(* IEC 61131-3 sources: Test002/ConveyorBelt/Class/SafetyBaseFSoE (part 5) *)

    end_if;

    //write to hardware from other module received SDO
    if ( ui_cnt_SDOInputBuffer > 0 ) & p_SDOInputBuffer then

      //set pointer to first SDO in the SDO list
      p_SDO_act   := p_SDOInputBuffer$^SDOHeader;

      //calculate length of SDO (CRC + data length)
      us_SDO_length := sizeof (SDOHeader.StdHeader.CRC) + p_SDO_act^.StdHeader.Len;

      //check, if buffer is empty
      if ( p_Handle_SDO_Write^.us_Status = SAFETY_SDO_NO_DATA ) then

#ifdef SAFETY_PROTOCOL_ANALYZER_ACTIVATED
  RecordFrame(p_SDO_act$^DINT, 1);
#endif

        //copy SDO into write-buffer
        ToStdLib.MemCpy(dest := #p_Handle_SDO_Write^.SDOStructure, source := p_SDO_act, size := us_SDO_length);

        //mark SDO data as valid
        p_Handle_SDO_Write^.us_Status := SAFETY_SDO_DATA_VALID;

        //decrement amount of SDOs
        ui_cnt_SDOInputBuffer -= 1;

        //if there is at least 1 SDO left, copy the remaining memory over the actual SDO
        if ( ui_cnt_SDOInputBuffer > 0 ) then

          //remove first entry in the SDO list
          _memmove(p_SDOInputBuffer, (p_SDOInputBuffer + SBF_SDO_MAX_LENGTH), (ui_cnt_SDOInputBuffer * SBF_SDO_MAX_LENGTH));
        end_if;
      end_if;
    end_if;

    if (b_ManagerInitialisationFinished = TRUE) & ( SafetyState <> _ReinitConfig ) & ( p_Handle_SDO_Write^.us_Status = SAFETY_SDO_NO_DATA ) then

      // priority request before checking the scheduler
      // if the channel is free and we have a command request for the flexible constellation node => send the command
      if (LastRequest = _NoOpenRequest) & (sFlexCon.FoundNodeInConfig) & (sFlexCon.CommandRequest) then

        StandardRequest.SDOHeader.CRC  := 0;                               // CRC is always 0 in Std communication
        StandardRequest.SDOHeader.Cmd  := SBF_SDO_COMMAND_WRITE;           // read command
        StandardRequest.SDOHeader.Typ  := SDO_STD;                         // standard frame type
        StandardRequest.SDOHeader.SeqNr:= StandardSeqNr OR 16#80;          // sequence number
        StandardRequest.SDOHeader.Len  := 4 + 4 + 1 + sizeof(UDINT);       // header + destination address + length of data + size of data
        StandardRequest.aData[0]$UDINT := SBF_SDO_ADDRESS_FLEX_CON_NODE;   // address of the flex con data
        StandardRequest.aData[4]       := sizeof(UDINT);                   // length of data
        StandardRequest.aData[5]$UDINT := sFlexCon.CommandRequest;     // new command

        // reset marker to detect new commands
        sFlexCon.CommandRequest := 0;

        LastRequest := _WriteFlexConCommand;

        //copy SDO into write-buffer
        ToStdLib.MemCpy(dest := #p_Handle_SDO_Write^.SDOStructure, source := #StandardRequest, size := (sizeof(SDOHeader.StdHeader.CRC) + StandardRequest.SDOHeader.Len));

        //mark SDO data as valid
        p_Handle_SDO_Write^.us_Status := SAFETY_SDO_DATA_VALID;

        if ( pISafety^.udVersion >= 16#1001 ) then
          SAFETY_iPushSafetyTask();
        end_if;

      end_if;

      // Start of scheduler; we need to share the time between reading, writing and diagnosis
      us_UnsafeSchedulerRun := 0;

      // number of steps in total minus 1, because the SetBusReady doesn't count here since it's not part of the rotation
      SchedulerStepNo := 10;

      // Check actions until we find somthing we need to do
      // all x (SchedulerStepNo) action-steps must be walked through during one cycle to make sure new data is fetched as fast as possible
      // SetBusReady is an exception: this step is only performed once on bootup!
      while (us_UnsafeSchedulerRun < SchedulerStepNo) & (LastRequest = _NoOpenRequest) do
        us_UnsafeSchedulerRun += 1;
        ud_UnsafeTimeoutCounter := 0; //No active request: we can reset the timeout-counter
        case UnsafeScheduler of
//**********************************************************************************************************************************************************
          UnsafeSchedulerSetBusReady:  // this step is excluded from the rotation (set at startup, on disconnect or quit error)

            case us_SetBusReadyState of

            //-------------------------------------------------------------------------------------------------------------
              WaitPDOsSyncron:

                EverythingSynchron := TRUE;

                // it's possible that all PDOs are coming from a different domain, then we have no inputbuffer
                if ui_cnt_PDOInputBuffer then
                  p_PDOInBufferAct := #aPDOInputBuffer[0];
                  for i := 0 to (ui_cnt_PDOInputBuffer-1) do
                    if p_PDOInBufferAct^.b_TimeSynchron = FALSE then
                      // we're still not synchron with this module. if it's optional it is probably not connected
                      if p_PDOInBufferAct^.b_IsOptional then
                        if (ops.tAbsolute - ud_OptionalTimeoutStart) <= SBF_OPTIONAL_MODULE_SYNC_TIMEOUT then
                          // if timeout not exceeded => not sychron (otherwise the variable will stay on it's old value)
                          EverythingSynchron := FALSE;
                          exit;
                        else
                          TRACE("Synchronisation timeout for optional module exceeded => assume it's synchon.");
                        end_if;
                      else
                        EverythingSynchron := FALSE;
                        exit;
                      end_if;
                    end_if;

                    p_PDOInBufferAct +=  sizeof(PDOInputBuffer);
                  end_for;

                  if EverythingSynchron & (ModuleSyncNo > 0) then
                    ModuleSyncNo -= 1;

#ifdef SAFETY_DEBUG_LOGGING_ACTIVATED
//                  case ud_MyModuleID of
//                    CSCP01x_ID:
//                      TRACE("ModuleSyncNo wurde dekrementiert von: CSCP.");
//
//                    CSDI16x_ID:
//                      TRACE("ModuleSyncNo wurde dekrementiert von: CSDI.");
//
//                    CSTO08x_ID:
//                      TRACE("ModuleSyncNo wurde dekrementiert von: CSTO.");
//                  end_case;
#endif
                end_if;
#ifdef SAFETY_DEBUG_LOGGING_ACTIVATED
//              elsif EverythingSynchron then
//                  case ud_MyModuleID of
//                    CSCP01x_ID:
//                      TRACE("ModuleSyncNo wurde nicht verändert von: CSCP.");
//
//                    CSDI16x_ID:
//                      TRACE("ModuleSyncNo wurde nicht verändert von: CSDI.");
//
//                    CSTO08x_ID:
//                      TRACE("ModuleSyncNo wurde nicht verändert von: CSTO.");
//                  end_case;
#endif
                end_if;

                if EverythingSynchron then
                  us_SetBusReadyState := WaitAllModulesSyncron;
                end_if;

            //-------------------------------------------------------------------------------------------------------------
              WaitAllModulesSyncron:
                // wait for other modules to be synchron with each other
                if (ModuleSyncNo = 0) & b_ManagerInitialisationFinished then
                  us_SetBusReadyState := SendSetBusReady;
                end_if;

            //-------------------------------------------------------------------------------------------------------------
              SendSetBusReady:
                // send the bus-ready command
                SDORequestBuffer.StdHeader.CRC  := 0;                                                   // CRC is always 0 in Std communication
                SDORequestBuffer.StdHeader.Cmd  := SBF_SDO_COMMAND_SET_BUS_READY;                        // set bus ready command
                SDORequestBuffer.StdHeader.Typ  := SDO_STD;                                             // standard frame type
                SDORequestBuffer.StdHeader.SeqNr:= StandardSeqNr OR 16#80;                              // sequence number
                SDORequestBuffer.StdHeader.Len  := 4;                                                   // header

                LastRequest := _SetBusReady;

#ifdef SAFETY_PROTOCOL_ANALYZER_ACTIVATED
  RecordFrame((#SDORequestBuffer)$^DINT, 1);
#endif

                //copy SDO into write-buffer
                ToStdLib.MemCpy(dest := #p_Handle_SDO_Write^.SDOStructure, source := #SDORequestBuffer, size := (sizeof(SDOHeader.StdHeader.CRC) + SDORequestBuffer.StdHeader.Len));

                //mark SDO data as valid
                p_Handle_SDO_Write^.us_Status := SAFETY_SDO_DATA_VALID;

                if ( pISafety^.udVersion >= 16#1001 ) then
                  SAFETY_iPushSafetyTask();
                end_if;

            //-------------------------------------------------------------------------------------------------------------
              SetBusReadyFinished:
                // all ok, nothing to do here

            end_case;
            us_UnsafeSchedulerRun := 16#FF; //make sure we don't repeat the while-loop until we have sent the bus-ready command

//**********************************************************************************************************************************************************
          UnsafeSchedulerGetDiagVars:

            //check, if buffer is empty and we got some unsafe data to get/set and crc check is finished
            if (DiagVars.SavingLogSSW = GetLogFileBlocks) then

              // check if more than blocksize to get
              if DiagVars.LogMemToGet > SBF_LOG_DATA_BLOCK_SIZE then
                // get a complete block
                DiagVars.BytesToGet := SBF_LOG_DATA_BLOCK_SIZE;
              else
                // get only the last bytes
                DiagVars.BytesToGet := DiagVars.LogMemToGet$USINT;
              end_if;

              StandardRequest.SDOHeader.Cmd   := SBF_SDO_COMMAND_READ;                         // read command
              StandardRequest.SDOHeader.Typ   := SDO_STD;                                     // standard frame type
              StandardRequest.SDOHeader.SeqNr := StandardSeqNr OR 16#80;                      // sequence number is in special area
              StandardRequest.SDOHeader.Len   := 4 + 4 + 1;                                   // header + destination address + length of data
              StandardRequest.aData[0]$UDINT  := DiagVars.ReadBaseAdr + (DiagVars.LogHeader.LogMemSize - DiagVars.LogMemToGet);// destination address
              StandardRequest.aData[4]        := DiagVars.BytesToGet$USINT;                   // length of data

              LastRequest := _ReadData;

#ifdef SAFETY_PROTOCOL_ANALYZER_ACTIVATED
  RecordFrame((#StandardRequest)$^DINT, 1);
#endif

              //copy SDO into write-buffer
              ToStdLib.MemCpy(dest := #p_Handle_SDO_Write^.SDOStructure, source := #StandardRequest, size := (sizeof(SDOHeader.StdHeader.CRC) + StandardRequest.SDOHeader.Len));

              //mark SDO data as valid
              p_Handle_SDO_Write^.us_Status := SAFETY_SDO_DATA_VALID;

              if ( pISafety^.udVersion >= 16#1001 ) then
                SAFETY_iPushSafetyTask();
              end_if;
            else
              UnsafeScheduler := UnsafeSchedulerNonPriorData;
            end_if;

//**********************************************************************************************************************************************************
          UnsafeSchedulerNonPriorData:

            // every 5 secs check for a new safety project inside the cpu
            if b_CheckCRC & ((ops.tAbsolute - ud_LastCrcCheck) > SBF_CRC_CHECK_TIME ) then

              SDORequestBuffer.StdHeader.CRC  := 0;                                                         // CRC is always 0 in Std communication
              SDORequestBuffer.StdHeader.Cmd  := SBF_SDO_COMMAND_READ;                                       // read command
              SDORequestBuffer.StdHeader.Typ  := SDO_STD;                                                   // standard frame type
              SDORequestBuffer.StdHeader.SeqNr:= StandardSeqNr OR 16#80;                                    // sequence number
              SDORequestBuffer.StdHeader.Len  := 4 + 4 + 1;                                                 // header + destination address + length of data
              SDORequestBuffer.ud_Address     := SBF_SDO_ADDRESS_CONFIG_DATA + SBF_SDO_OFFSET_CONFIG_CRC_ALL; // address of crc
              SDORequestBuffer.us_Length      := 4;                                                         // length of crc

              LastRequest := _GetCRC;

#ifdef SAFETY_PROTOCOL_ANALYZER_ACTIVATED
  RecordFrame((#SDORequestBuffer)$^DINT, 1);
#endif

              //copy SDO into write-buffer
              ToStdLib.MemCpy(dest := #p_Handle_SDO_Write^.SDOStructure, source := #SDORequestBuffer, size := (sizeof(SDOHeader.StdHeader.CRC) + SDORequestBuffer.StdHeader.Len));

              //mark SDO data as valid
              p_Handle_SDO_Write^.us_Status := SAFETY_SDO_DATA_VALID;

              if ( pISafety^.udVersion >= 16#1001 ) then
                SAFETY_iPushSafetyTask();
              end_if;

              ud_LastCrcCheck := ops.tAbsolute;

            // every 5 seconds write system time of plc to scp
            elsif b_SetSysTime & ((ops.tAbsolute - ud_LastSetSysTime) > SBF_SYSTIME_SET_TIME ) then

              if (LastRequest = _NoOpenRequest) & (p_Handle_SDO_Write^.us_Status = SAFETY_SDO_NO_DATA) then
                StandardRequest.SDOHeader.CRC  := 0;                               // CRC is always 0 in Std communication
                StandardRequest.SDOHeader.Cmd  := SBF_SDO_COMMAND_WRITE;           // read command
                StandardRequest.SDOHeader.Typ  := SDO_STD;                         // standard frame type
                StandardRequest.SDOHeader.SeqNr:= StandardSeqNr OR 16#80;          // sequence number
                StandardRequest.SDOHeader.Len  := 4 + 4 + 1 + sizeof(UDINT);       // header + destination address + length of data + size of data
                StandardRequest.aData[0]$UDINT := SBF_SDO_ADDRESS_FW_SYSTIME;      // address of system time safety firmware
                StandardRequest.aData[4]       := sizeof(UDINT);                   // length of data
                StandardRequest.aData[5]$UDINT := ToSigCLib.UnixTimeStampGet();    // system time of plc as unix timestamp

                LastRequest := _WriteSysTime;

                //copy SDO into write-buffer
                ToStdLib.MemCpy(dest := #p_Handle_SDO_Write^.SDOStructure, source := #StandardRequest, size := (sizeof(SDOHeader.StdHeader.CRC) + StandardRequest.SDOHeader.Len));

                //mark SDO data as valid
                p_Handle_SDO_Write^.us_Status := SAFETY_SDO_DATA_VALID;

                if ( pISafety^.udVersion >= 16#1001 ) then
                  SAFETY_iPushSafetyTask();
                end_if;

                ud_LastSetSysTime := ops.tAbsolute;
              end_if;

            else
              if RunState then
                // in operational also get unsave-variables
                UnsafeScheduler := UnsafeSchedulerWriteData;
              else
                // not operational, we must skip the unsave vars
                UnsafeScheduler := UnsafeSchedulerDiagState;
                us_UnsafeSchedulerRun += 2;
              end_if;
            end_if;

//**********************************************************************************************************************************************************
          UnsafeSchedulerWriteData:

            if IsOptimizedCPU() then
              if ui_CntUnsafeInputs then
                // if we have finished checking through all variables the last time => check from beginning (otherwise the pointer is on the element where we have to continue)
                if pUnsafeInElement = NIL then
                  pUnsafeInElement := p_UnsafeInputsTable;
                end_if;

                // we check if we have to write any of the unsafe input variables (only until our message is full)
                UnsafeWrPackageNo := 0;
                BDINTWriteVars := 0; // limit number of bdint write variables to 3 to ensure constant load of firmware
                while pUnsafeInElement & (UnsafeWrPackageNo < SBF_MAX_UNSAFE_WRITE_PACKAGES) & (BDINTWriteVars < SBF_MAX_UNSAFE_BDINTS_PER_WRITE) do

                  // we have to check if we add this one
                  GotNewUnsafeValue := FALSE;

                  // if the type is normal we can read the actual value from the server
                  if pUnsafeInElement^.UnsafeType = NormalUnsafe then
                    // check if pointer to server is valid
                    if pUnsafeInElement^.ud_Thisp then
                      // get the actual value from the server
                      TmpVal := RD((pUnsafeInElement^.ud_Thisp)$^void);

                      // we remember to update this if it's necessary
                      GotNewUnsafeValue := TRUE;
                    else
                      if bd_LogOnceMarker.NoThisForUnsafeIn = FALSE then
                        bd_LogOnceMarker.NoThisForUnsafeIn := TRUE;
                        LogError("@0269 (SafetyBaseFSoE::CyWork) [SL] No thispointer available for Server of local unsafe input variable.");
                      end_if;
                    end_if;
                  elsif pUnsafeInElement^.UnsafeType = ExternalInput then
                    // check if we already have a valid value there
                    if pUnsafeInElement^.b_IsValid then
                      // get the actual value from the element
                      TmpVal := pUnsafeInElement^.sd_NewValue4External;

                      // we remember to update this if it's necessary
                      GotNewUnsafeValue := TRUE;
                    end_if;
                  else
                    if bd_LogOnceMarker.WrongUnsafeVarType = FALSE then
                      bd_LogOnceMarker.WrongUnsafeVarType := TRUE;
                      LogError("@026A (SafetyBaseFSoE::CyWork) [SL] Wrong unsafe variable type in unsafe input list.");
                    end_if;
                  end_if;

                  // if we have a new valid unsafe value => check if we have to send it
                  if GotNewUnsafeValue then
                    // if it hasn't been sent yet
                    if (pUnsafeInElement^.b_AlreadyTransmitted = FALSE) then
                      // remember that we sent this already
                      pUnsafeInElement^.b_AlreadyTransmitted := TRUE;

                      // add this one
                      AddUnsafePackage := TRUE;
                    elsif TmpVal <> pUnsafeInElement^.sd_OldValue then
                      // if there were any changes on this value

                      // add this one
                      AddUnsafePackage := TRUE;
                    else
                      // don't add this one
                      AddUnsafePackage := FALSE;
                    end_if;

                    // if it is ready to be added => add it to send buffer
                    if AddUnsafePackage then
                      // add a package to send
                      aUnsafeWrPackages[UnsafeWrPackageNo].ud_Address := pUnsafeInElement^.ud_Address;
                      aUnsafeWrPackages[UnsafeWrPackageNo].Value      := TmpVal;
                      UnsafeWrPackageNo += 1;

                      // if it has a bitmask it's an unsafe bdint input variable
                      if pUnsafeInElement^.BitMask then
                        BDINTWriteVars += 1;
                      end_if;

                      // remember the actual as old value
                      pUnsafeInElement^.sd_OldValue := TmpVal;
                    end_if;
                  end_if;

                  pUnsafeInElement := pUnsafeInElement^.pNext;
                end_while;

                if UnsafeWrPackageNo then
                  DataLen := UnsafeWrPackageNo * sizeof(UnsafeWritePackage);

                  StandardRequest.SDOHeader.Cmd                 := SBF_SDO_COMMAND_WRITE_VALUES;    // write values command
                  StandardRequest.SDOHeader.Typ                 := SDO_STD;                        // standard frame type
                  StandardRequest.SDOHeader.SeqNr               := StandardSeqNr OR 16#80;         // sequence number is in special area
                  StandardRequest.SDOHeader.Len                 := 4 + 4 + 1 + DataLen;            // header + destination address + length of data + data
                  StandardRequest.aData[0]                      := UnsafeWrPackageNo;              // number of packages
                  StandardRequest.aData[1]$UnsafeWritePackages  := aUnsafeWrPackages;              // packages

                  LastRequest := _WriteValues;

#ifdef SAFETY_PROTOCOL_ANALYZER_ACTIVATED
  RecordFrame((#StandardRequest)$^DINT, 1);
#endif

                  //copy SDO into write-buffer
                  ToStdLib.MemCpy(dest := #p_Handle_SDO_Write^.SDOStructure, source := #StandardRequest, size := (sizeof(SDOHeader.StdHeader.CRC) + StandardRequest.SDOHeader.Len));

                  //mark SDO data as valid
                  p_Handle_SDO_Write^.us_Status := SAFETY_SDO_DATA_VALID;

                  if ( pISafety^.udVersion >= 16#1001 ) then
                    SAFETY_iPushSafetyTask();
                  end_if;
                else
                  UnsafeScheduler := UnsafeSchedulerReadData;
                end_if;
              else
                UnsafeScheduler := UnsafeSchedulerReadData;
              end_if;
            else
              // on CSCP011 the SDO_COMMAND_WRITE_VALUES didn't exist
              if ui_CntUnsafeInputs & WriteFramesNeeded then
                // if writing is not active, check if it's necessary to activate it
                if (UnsafeWritingActive = FALSE) then
                  pUnsafeInElement := p_UnsafeInputsTable;

                  for i := 0 to (ui_CntUnsafeInputs - 1) do
                    if pUnsafeInElement^.ud_Thisp then
                      sd_retval := RD((pUnsafeInElement^.ud_Thisp)$^void);        // data
                      if pUnsafeInElement^.sd_OldValue <> sd_retval then
                        UnsafeWritingActive := TRUE;
                        pUnsafeInElement^.sd_OldValue := sd_retval;
                      end_if;
                    end_if;
                    pUnsafeInElement += sizeof(UnsafeIORoutingElement);
                  end_for;
                end_if;

                // check if writing is already active
                if UnsafeWritingActive then
                  // pointer to the right unsafe input
                  pUnsafeInElement := p_UnsafeInputsTable + (UnsafeWriteTransNr * MaxVarsPerWritePackage * sizeof(UnsafeIORoutingElement));

                  // get length of data we write
                  if (UnsafeWriteTransNr < (WriteFramesNeeded-1)) | ((ui_CntUnsafeInputs MOD MaxVarsPerWritePackage) = 0) then
                    DataLen := MaxVarsPerWritePackage * sizeof(DINT);
                  else
                    DataLen := (ui_CntUnsafeInputs MOD MaxVarsPerWritePackage)$USINT * sizeof(DINT);
                  end_if;

                  StandardRequest.SDOHeader.Cmd   := SBF_SDO_COMMAND_WRITE;                        // write command
                  StandardRequest.SDOHeader.Typ   := SDO_STD;                                     // standard frame type
                  StandardRequest.SDOHeader.SeqNr := StandardSeqNr OR 16#80;                      // sequence number is in special area
                  StandardRequest.SDOHeader.Len   := 4 + 4 + 1 + DataLen;                         // header + destination address + length of data + data
                  StandardRequest.aData[0]$UDINT  := pUnsafeInElement^.ud_Address;                // destination address
                  StandardRequest.aData[4]        := DataLen;                                     // length of data

                  // depending on length we do different number of server read-methods to get the data we write
                  for i := 0 to (DataLen/sizeof(DINT)) - 1 do
                    if pUnsafeInElement^.ud_Thisp then
                      StandardRequest.aData[5 + (i * sizeof(DINT))]$DINT := pUnsafeInElement^.sd_OldValue;
                    else
                      // this server doesn't exist in lasal => always send 0
                      StandardRequest.aData[5 + (i * sizeof(DINT))]$DINT := 0;
                    end_if;

                    pUnsafeInElement += sizeof(UnsafeIORoutingElement);
                  end_for;

                  LastRequest := _WriteValues;

#ifdef SAFETY_PROTOCOL_ANALYZER_ACTIVATED
  RecordFrame((#StandardRequest)$^DINT, 1);
#endif

                  //copy SDO into write-buffer
                  ToStdLib.MemCpy(dest := #p_Handle_SDO_Write^.SDOStructure, source := #StandardRequest, size := (sizeof(SDOHeader.StdHeader.CRC) + StandardRequest.SDOHeader.Len));

                  //mark SDO data as valid
                  p_Handle_SDO_Write^.us_Status := SAFETY_SDO_DATA_VALID;

                  if ( pISafety^.udVersion >= 16#1001 ) then
                    SAFETY_iPushSafetyTask();
                  end_if;
                else
                  UnsafeScheduler := UnsafeSchedulerReadData;
                end_if;
              else
                UnsafeScheduler := UnsafeSchedulerReadData;
              end_if;
            end_if;

//**********************************************************************************************************************************************************
          UnsafeSchedulerReadData:

            if ui_CntUnsafeOutputs & ReadFramesNeeded then
              //check, if buffer is empty and we got some unsafe data to get/set and crc check is finished
              if (UnsafeReadTransNr < ReadFramesNeeded) //then
               & ( ((UnsafeReadTransNr = 0) & ( ops.tAbsolute - LastUnsafeUpdate > ud_ServerUpdateTime ) ) | (UnsafeReadTransNr <> 0) )then
                // here we request directly the unsafe IOs

                // sequence number is in special area
                StandardRequest.SDOHeader.SeqNr := StandardSeqNr OR 16#80;

                // we get an output
                pUnsafeOutElement := p_UnsafeOutputsTable + (UnsafeReadTransNr * MaxVarsPerReadPackage * sizeof(UnsafeIORoutingElement));

                // get length of data we read
                if (UnsafeReadTransNr < (ReadFramesNeeded - 1)) | ((ui_CntUnsafeOutputs MOD MaxVarsPerReadPackage) = 0) then
                  UnsafeRdPackageNo := MaxVarsPerReadPackage;
                else
                  UnsafeRdPackageNo := (ui_CntUnsafeOutputs MOD MaxVarsPerReadPackage)$USINT;
                end_if;

                DataLen := UnsafeRdPackageNo * sizeof(DINT);

                // create buffer with addresses of values to read
                pHelpUnsafe := pUnsafeOutElement;
                for i := 0 to (UnsafeRdPackageNo-1) do
                  aUnsafeRdPackages[i] := pHelpUnsafe^.ud_Address;
                  pHelpUnsafe += sizeof(UnsafeIORoutingElement);
                end_for;

                StandardRequest.SDOHeader.Cmd               := SBF_SDO_COMMAND_READ_VALUES;                  // read values command
                StandardRequest.SDOHeader.Typ               := SDO_STD;                                     // standard frame type
                StandardRequest.SDOHeader.SeqNr             := StandardSeqNr OR 16#80;                      // sequence number is in special area
                StandardRequest.SDOHeader.Len               := 4 + 1 + DataLen;                             // header + size + length of data
                StandardRequest.aData[0]                    := UnsafeRdPackageNo;                           // number of values to get
                StandardRequest.aData[1]$UnsafeReadPackages := aUnsafeRdPackages;                           // read addresses

                LastRequest := _ReadValues;

#ifdef SAFETY_PROTOCOL_ANALYZER_ACTIVATED
  RecordFrame((#StandardRequest)$^DINT, 1);
#endif

                //copy SDO into write-buffer
                ToStdLib.MemCpy(dest := #p_Handle_SDO_Write^.SDOStructure, source := #StandardRequest, size := (sizeof(SDOHeader.StdHeader.CRC) + StandardRequest.SDOHeader.Len));

                //mark SDO data as valid
                p_Handle_SDO_Write^.us_Status := SAFETY_SDO_DATA_VALID;

                if ( pISafety^.udVersion >= 16#1001 ) then
                  SAFETY_iPushSafetyTask();
                end_if;

              elsif (UnsafeReadTransNr >= ReadFramesNeeded) then
                // We have finished all read data, go on with the next step
                UnsafeScheduler := UnsafeSchedulerDiagState;
                LastUnsafeUpdate := ops.tAbsolute;
                UnsafeReadTransNr := 0;
              else
                // time until read is not yet over - go on
                UnsafeScheduler := UnsafeSchedulerDiagState;
              end_if;
            else
              UnsafeScheduler := UnsafeSchedulerDiagState;
            end_if;

//**********************************************************************************************************************************************************
          UnsafeSchedulerDiagState:

            // get the diag state (on user demand)
            if DiagVars.UserWantsDiagState then

              // get state via SDO communication
              SDORequestBuffer.StdHeader.CRC  := 0;                                                   // CRC is always 0 in Std communication
              SDORequestBuffer.StdHeader.Cmd  := SBF_SDO_COMMAND_GET_STATE;                            // get-state command
              SDORequestBuffer.StdHeader.Typ  := SDO_STD;                                             // standard frame type
              SDORequestBuffer.StdHeader.SeqNr:= StandardSeqNr OR 16#80;                              // sequence number
              SDORequestBuffer.StdHeader.Len  := 4;                                                   // header
              SDORequestBuffer.ud_Address     := 0;
              SDORequestBuffer.us_Length      := 0;

              LastRequest := _DiagState;

#ifdef SAFETY_PROTOCOL_ANALYZER_ACTIVATED
  RecordFrame((#SDORequestBuffer)$^DINT, 1);
#endif

              //copy SDO into write-buffer
              ToStdLib.MemCpy(dest := #p_Handle_SDO_Write^.SDOStructure, source := #SDORequestBuffer, size := (sizeof(SDOHeader.StdHeader.CRC) + SDORequestBuffer.StdHeader.Len));

              //mark SDO data as valid
              p_Handle_SDO_Write^.us_Status := SAFETY_SDO_DATA_VALID;

              if ( pISafety^.udVersion >= 16#1001 ) then
                SAFETY_iPushSafetyTask();
              end_if;
            else
              UnsafeScheduler := UnsafeSchedulerDiagInfo;
            end_if;

//**********************************************************************************************************************************************************
            UnsafeSchedulerDiagInfo:

            // get the diag info (on user demand)
            if DiagVars.UserWantsDiagInfo then

              // get state via SDO communication
              StandardRequest.SDOHeader.CRC  := 0;                                                   // CRC is always 0 in Std communication
              StandardRequest.SDOHeader.Cmd  := SBF_SDO_COMMAND_GET_DIAG_INFO;                        // read command
              StandardRequest.SDOHeader.Typ  := SDO_STD;                                             // standard frame type
              StandardRequest.SDOHeader.SeqNr:= StandardSeqNr OR 16#80;                              // sequence number
              StandardRequest.SDOHeader.Len  := 4 + 1;                                               // header + µC-selection
              StandardRequest.aData[0] := DiagVars.ucChoiceDiagInfo;

              LastRequest := _DiagInfo;

#ifdef SAFETY_PROTOCOL_ANALYZER_ACTIVATED
  RecordFrame((#StandardRequest)$^DINT, 1);
#endif

              //copy SDO into write-buffer
              ToStdLib.MemCpy(dest := #p_Handle_SDO_Write^.SDOStructure, source := #StandardRequest, size := (sizeof(SDOHeader.StdHeader.CRC) + StandardRequest.SDOHeader.Len));

              //mark SDO data as valid
              p_Handle_SDO_Write^.us_Status := SAFETY_SDO_DATA_VALID;

              if ( pISafety^.udVersion >= 16#1001 ) then
                SAFETY_iPushSafetyTask();
              end_if;

            else

//              if SchedulerStepNo = 6 then
//                UnsafeScheduler := UnsafeSchedulerGetDiagVars;
//
//              elsif SchedulerStepNo = 7 then
//                UnsafeScheduler := UnsafeSchedulerGetRetryCounter;
//              end_if;
              UnsafeScheduler := UnsafeSchedulerGetRetryCounter;

            end_if;

//**********************************************************************************************************************************************************
          UnsafeSchedulerGetRetryCounter:

            //read out the retry counters every 10seconds
            if (b_RetryCounterAvailable) & (b_DisableSafetyRetryCnt = FALSE)
            & ((ops.tAbsolute - ud_RetryCntTimeMark) > SBF_RETRY_COUNTER_WAIT_TIME)  then

              SDORequestBuffer.StdHeader.CRC  := 0;                                                         // CRC is always 0 in Std communication
              SDORequestBuffer.StdHeader.Cmd  := SBF_SDO_COMMAND_READ;                                       // read command
              SDORequestBuffer.StdHeader.Typ  := SDO_STD;                                                   // standard frame type
              SDORequestBuffer.StdHeader.SeqNr:= StandardSeqNr OR 16#80;                                    // sequence number
              SDORequestBuffer.StdHeader.Len  := 4 + 4 + SBF_SDO_LENGTH_RETRY_COUNTER;                       // header + destination address + length of data
              SDORequestBuffer.ud_Address     := SBF_SDO_ADDRESS_RETRY_COUNTER;                              // address of retrycounter
              SDORequestBuffer.us_Length      := SBF_SDO_LENGTH_RETRY_COUNTER;                               // length of data

              LastRequest := _ReadRetryCounter;

#ifdef SAFETY_PROTOCOL_ANALYZER_ACTIVATED
  RecordFrame((#SDORequestBuffer)$^DINT, 1);
#endif

              //copy SDO into write-buffer
              ToStdLib.MemCpy(dest := #p_Handle_SDO_Write^.SDOStructure, source := #SDORequestBuffer, size := (sizeof(SDOHeader.StdHeader.CRC) + SDORequestBuffer.StdHeader.Len));

              //mark SDO data as valid
              p_Handle_SDO_Write^.us_Status := SAFETY_SDO_DATA_VALID;

              if ( pISafety^.udVersion >= 16#1001 ) then
                SAFETY_iPushSafetyTask();
              end_if;

              //reset timemark
              ud_RetryCntTimeMark := ops.tAbsolute;

            else
              UnsafeScheduler := UnsafeSchedulerChannelError;
            end_if;

//**********************************************************************************************************************************************************
          UnsafeSchedulerChannelError:

            if DiagVars.UserWantsErrorInfo  then
              SDORequestBuffer.StdHeader.CRC  := 0;                                                          // CRC is always 0 in Std communication
              SDORequestBuffer.StdHeader.Cmd  := SBF_SDO_COMMAND_READ;                                       // read command
              SDORequestBuffer.StdHeader.Typ  := SDO_STD;                                                    // standard frame type
              SDORequestBuffer.StdHeader.SeqNr:= StandardSeqNr OR 16#80;                                     // sequence number
              SDORequestBuffer.StdHeader.Len  := 4 + 4 + 1;                                                  // header + destination address + length of data
              SDORequestBuffer.ud_Address     := SBF_SDO_ADDRESS_ERROR_MEM;                                  // address of error memory
              SDORequestBuffer.us_Length      := SBF_SDO_LENGTH_ERROR_MESSAGE;                               // length of data (first byte contains number of following values + number of channels)

              if remainingPacketlength <> 0 then
                // set offset if more than one package
                SDORequestBuffer.ud_Address     := (SBF_SDO_ADDRESS_ERROR_MEM + actoffset);                  // address of error memory
                // set new length for next package
                if remainingPacketlength > SBF_SDO_LENGTH_ERROR_MESSAGE then
                  SDORequestBuffer.us_Length      := SBF_SDO_LENGTH_ERROR_MESSAGE;
                else
                  SDORequestBuffer.us_Length      := remainingPacketlength$USINT;
                end_if;
              end_if;

              LastRequest := _ErrorChannelInfo;

#ifdef SAFETY_PROTOCOL_ANALYZER_ACTIVATED
RecordFrame((#SDORequestBuffer)$^DINT, 1);
#endif

              //copy SDO into write-buffer
              ToStdLib.MemCpy(dest := #p_Handle_SDO_Write^.SDOStructure, source := #SDORequestBuffer, size := (sizeof(SDOHeader.StdHeader.CRC) + SDORequestBuffer.StdHeader.Len));

              //mark SDO data as valid
              p_Handle_SDO_Write^.us_Status := SAFETY_SDO_DATA_VALID;

              if ( pISafety^.udVersion >= 16#1001 ) then
                SAFETY_iPushSafetyTask();
              end_if;

              //reset timemark
              ud_RetryCntTimeMark := ops.tAbsolute;

            else
              UnsafeScheduler := UnsafeSchedulerGetFlexConNodeState;
            end_if;

//**********************************************************************************************************************************************************
          UnsafeSchedulerGetFlexConNodeState:

            // if there is a flexible constellation in the configuration and also an object placed and connected, we check the state regularly
            if (sFlexCon.FoundNodeInConfig) & ((ops.tAbsolute - sFlexCon.ud_LastNodeStateTimeStamp) > SBF_FLEX_CON_STATE_CHECK_TIME) then

              SDORequestBuffer.StdHeader.CRC  := 0;                                                         // CRC is always 0 in Std communication
              SDORequestBuffer.StdHeader.Cmd  := SBF_SDO_COMMAND_READ;                                      // read command
              SDORequestBuffer.StdHeader.Typ  := SDO_STD;                                                   // standard frame type
              SDORequestBuffer.StdHeader.SeqNr:= StandardSeqNr OR 16#80;                                    // sequence number
              SDORequestBuffer.StdHeader.Len  := 4 + 4 + sizeof(t_FlexConNodeState);                        // header + destination address + length of data
              SDORequestBuffer.ud_Address     := SBF_SDO_ADDRESS_FLEX_CON_NODE;                             // address of retrycounter
              SDORequestBuffer.us_Length      := sizeof(t_FlexConNodeState);                                // length of data

              LastRequest := _ReadFlexConNodeState;

#ifdef SAFETY_PROTOCOL_ANALYZER_ACTIVATED
  RecordFrame((#SDORequestBuffer)$^DINT, 1);
#endif

              //copy SDO into write-buffer
              ToStdLib.MemCpy(dest := #p_Handle_SDO_Write^.SDOStructure, source := #SDORequestBuffer, size := (sizeof(SDOHeader.StdHeader.CRC) + SDORequestBuffer.StdHeader.Len));

              //mark SDO data as valid
              p_Handle_SDO_Write^.us_Status := SAFETY_SDO_DATA_VALID;

              if ( pISafety^.udVersion >= 16#1001 ) then
                SAFETY_iPushSafetyTask();
              end_if;

              //reset timemark
              sFlexCon.ud_LastNodeStateTimeStamp := ops.tAbsolute;

            else
              UnsafeScheduler := UnsafeSchedulerGetFlexConHostState;
            end_if;

//**********************************************************************************************************************************************************
          UnsafeSchedulerGetFlexConHostState:

            // if there is a flexible constellation in the configuration and also an object placed and connected, we check the state regularly
            if (sFlexCon.FoundHostInConfig) & ((ops.tAbsolute - sFlexCon.ud_LastHostStateTimeStamp) > SBF_FLEX_CON_STATE_CHECK_TIME) then

              // calcuate max length
              us_SDO_length := SBF_SDO_MAX_LENGTH - (sizeof(SDOHeader) - sizeof(SDOHeader.SessId)) - sizeof(SDORespReadConfig.us_Returncode) - sizeof(SDORespReadConfig.us_Length);

              // if it's the first read of this run, read as much as possible (we don't know how many connections we have yet)
              if sFlexCon.LastHostState.CurrentReadOffset = 0 then
                // get maximum number of bytes
                DataLen := us_SDO_length;
              else
                // if we still need more or equal to max size
                if sFlexCon.LastHostState.BytesMissing >= us_SDO_length then
                  // get maximum number of bytes
                  DataLen := us_SDO_length;
                else
                  // otherwise it's the last package, so get the rest that is missing
                  DataLen := sFlexCon.LastHostState.BytesMissing$USINT;
                end_if;
              end_if;

              SDORequestBuffer.StdHeader.CRC  := 0;                                                                         // CRC is always 0 in Std communication
              SDORequestBuffer.StdHeader.Cmd  := SBF_SDO_COMMAND_READ;                                                      // read command
              SDORequestBuffer.StdHeader.Typ  := SDO_STD;                                                                   // standard frame type
              SDORequestBuffer.StdHeader.SeqNr:= StandardSeqNr OR 16#80;                                                    // sequence number
              SDORequestBuffer.StdHeader.Len  := 4 + 4 + sizeof(HDINT);                                                     // header + destination address + length of data
              SDORequestBuffer.ud_Address     := SBF_SDO_ADDRESS_FLEX_CON_HOST + sFlexCon.LastHostState.CurrentReadOffset;  // address of retrycounter
              SDORequestBuffer.us_Length      := DataLen;                                                                   // length of data

              // remember the length to check it when we receive the answer
              sFlexCon.LastHostState.LastRequestedLength := DataLen;

              LastRequest := _ReadFlexConHostState;

#ifdef SAFETY_PROTOCOL_ANALYZER_ACTIVATED
  RecordFrame((#SDORequestBuffer)$^DINT, 1);
#endif

              //copy SDO into write-buffer
              ToStdLib.MemCpy(dest := #p_Handle_SDO_Write^.SDOStructure, source := #SDORequestBuffer, size := (sizeof(SDOHeader.StdHeader.CRC) + SDORequestBuffer.StdHeader.Len));

              //mark SDO data as valid
              p_Handle_SDO_Write^.us_Status := SAFETY_SDO_DATA_VALID;

              if ( pISafety^.udVersion >= 16#1001 ) then
                SAFETY_iPushSafetyTask();
              end_if;

            else
              UnsafeScheduler := UnsafeSchedulerGetDiagVars;
            end_if;

//**********************************************************************************************************************************************************
        else
          if bd_LogOnceMarker.InvalidSchedulerState = FALSE then
            bd_LogOnceMarker.InvalidSchedulerState := TRUE;
            LogError("@026B (SafetyBaseFSoE::CyWork) [SL] Undefined Scheduler-State.");
          end_if;
        end_case;
      end_while;
    end_if;
  end_if;

  // at the first run we write all variables independent of any changes
  if RunState > OldRunState then
    SendAllUnsafeValues();
  end_if;
  OldRunState := RunState;

  state := READY;

//============================ Profiler start======================================================
#ifdef  DM_Profiler
  StopTimeMeasurement(usMode := DMTIME_CY);
#endif
//============================ Profiler end========================================================
END_FUNCTION

FUNCTION VIRTUAL SafetyBaseFSoE::GetConfiguration

END_FUNCTION

FUNCTION VIRTUAL SafetyBaseFSoE::SetSafetyState
  VAR_INPUT
    NewState 	: SafetyConfigStateType;
  END_VAR

  // use it locally => can also be forwarded in derivation
  SafetyState := NewState;

END_FUNCTION

FUNCTION VIRTUAL SafetyBaseFSoE::RefreshAsySrv
  // derive this
END_FUNCTION

FUNCTION VIRTUAL SafetyBaseFSoE::SetRetryCounter

  SafetyRetryCounter := -1;

END_FUNCTION

FUNCTION SafetyBaseFSoE::IsInCache
  VAR_INPUT
    ud_Address 	: UDINT;
    us_Length 	: USINT;
  END_VAR
  VAR_OUTPUT
    ItsInside 	: BOOL;
  END_VAR

  if CachedSize &
     (ud_Address >= CachedAddr) &
     ((ud_Address + us_Length) <= (CachedAddr + CachedSize)) then
    ItsInside := TRUE;
  else
    ItsInside := FALSE;
  end_if;

END_FUNCTION

FUNCTION SafetyBaseFSoE::AddToCache
  VAR_INPUT
    p_SDORequestBuffer 	: ^SDORequReadConfig;
    p_SDOResponseBuffer 	: ^SDORespReadConfig;
  END_VAR

  if p_SDORequestBuffer^.us_Length then
    CachedAddr := p_SDORequestBuffer^.ud_Address;
    CachedSize := p_SDORequestBuffer^.us_Length;
    _memcpy(ptr1:=#Cache, ptr2:=#p_SDOResponseBuffer^.ud_Data, cntr:=p_SDORequestBuffer^.us_Length);
  end_if;

END_FUNCTION

FUNCTION SafetyBaseFSoE::GetFSoEConnectionInfos
  VAR_INPUT
    p_SDORequestBuffer 	: ^SafetyBaseFSoE::SDORequReadConfig;
    p_SDOResponseBuffer 	: ^SafetyBaseFSoE::SDORespReadConfig;
  END_VAR
  VAR
    Address         : UDINT;
    Size            : USINT;
    sd_retval       : DINT;
    i               : UDINT;
    pActConnection  : ^t_FSoEConnectionDetails;
    TempRoutingInfo : t_FSoERoutingInfoElement;
    NextAddress     : UDINT;
  END_VAR

  // free the list if there is still one
  FreeFSoEConnectionInfos();

  // check if we already got the info:
  if ConnectionInfos.ConnectionNo | ConnectionInfos.pFirstConnection then
    LogError("@0280 (SafetyBaseFSoE::GetFSoEConnectionInfos) List already exists! May not have been resetted correctly!");
    return;
  end_if;

//*****************************************************************************
//** CONNECTION STATE INFO                                                   **
//*****************************************************************************

  // get number of connections
  Address := SBF_SDO_ADDRESS_FSOE_CONN_STATE;
  Size    := 2;

  //send request and receive data
  sd_retval := SDOReadCfgRequ ( p_SDORequestBuffer  := p_SDORequestBuffer
                              , p_SDOResponseBuffer := p_SDOResponseBuffer
                              , ud_Address          := Address
                              , us_Length           := Size
                              );

  //no response
  if ( sd_retval <> 0 ) then
    LogError("@0281 (SafetyBaseFSoE::GetFSoEConnectionInfos) Config Read Error: Error reading number of connections.");
    return;
  end_if;

  ConnectionInfos.ConnectionNo := p_SDOResponseBuffer^.ud_Data$UINT;

  if ConnectionInfos.ConnectionNo = 0 then
    // no connections available
    return;
  end_if;

  // allocate memory for the connections
  ConnectionInfos.pFirstConnection$pVoid := ToStdLib.Malloc(size:= ConnectionInfos.ConnectionNo * sizeof(t_FSoEConnectionDetails));

  if ConnectionInfos.pFirstConnection = NIL then
    LogError("@0282 (SafetyBaseFSoE::GetFSoEConnectionInfos) Config Read Error: Failed to allocate memory for FSoE connection details.");
    return;
  end_if;

  // reset memory (also resets pNext although we are not using a linked list here)
  _memset(dest:=ConnectionInfos.pFirstConnection, usByte:=0, cntr:= ConnectionInfos.ConnectionNo * sizeof(t_FSoEConnectionDetails));

  Address += Size;
  Size    := 1;

  pActConnection := ConnectionInfos.pFirstConnection;

  // get connection states
  for i := 0 to ConnectionInfos.ConnectionNo-1 do
    // get state of connection

    //send request and receive data
    sd_retval := SDOReadCfgRequ ( p_SDORequestBuffer  := p_SDORequestBuffer
                                , p_SDOResponseBuffer := p_SDOResponseBuffer
                                , ud_Address          := Address
                                , us_Length           := Size
                                );

    //no response
    if ( sd_retval <> 0 ) then
      LogError("@0283 (SafetyBaseFSoE::GetFSoEConnectionInfos) Config Read Error: Error reading connection state.");
      return;
    end_if;

    // get connection state
    pActConnection^.ConnectionState := (p_SDOResponseBuffer^.ud_Data$USINT AND 2#0111)$t_FSoEConnectionState;

    // get info if the module is master or slave at this connection
    pActConnection^.Flags.IsMaster  := (p_SDOResponseBuffer^.ud_Data$USINT AND 2#1000) <> 0;

    // save safety number
    pActConnection^.OwnerSafetyNbr  := SafetyNumber;

    // for easier debugging we set the correct next pointers
    if i = ConnectionInfos.ConnectionNo-1 then
      pActConnection^.pNext := NIL;
    else
      pActConnection^.pNext := pActConnection + sizeof(t_FSoEConnectionDetails);
    end_if;

    pActConnection                  += sizeof(t_FSoEConnectionDetails);
    Address                         += Size;
  end_for;

//*****************************************************************************
//** ROUTING INFO                                                            **
//*****************************************************************************

  // get number of connections
  Address := SBF_SDO_ADDRESS_FSOE_ROUTING_INFO;
  Size    := 2;

  //send request and receive data
  sd_retval := SDOReadCfgRequ ( p_SDORequestBuffer  := p_SDORequestBuffer
                              , p_SDOResponseBuffer := p_SDOResponseBuffer
                              , ud_Address          := Address
                              , us_Length           := Size
                              );

  //no response
  if ( sd_retval <> 0 ) then
    LogError("@0281 (SafetyBaseFSoE::GetFSoEConnectionInfos) Config Read Error: Error reading number of connections.");
    return;
  end_if;

  // check if it's the same number
  if ConnectionInfos.ConnectionNo <> p_SDOResponseBuffer^.ud_Data$UINT then
    LogError("@0285 (SafetyBaseFSoE::GetFSoEConnectionInfos) Config Read Error: Number of connections does not match (case 1).");
    return;
  end_if;

  Address += Size;
  Size    := sizeof(t_FSoERoutingInfoElement);

  pActConnection := ConnectionInfos.pFirstConnection;

  // get connection states
  for i := 0 to ConnectionInfos.ConnectionNo-1 do
    // get routing info of connections

    //send request and receive data
    sd_retval := SDOReadCfgRequ ( p_SDORequestBuffer  := p_SDORequestBuffer
                                , p_SDOResponseBuffer := p_SDOResponseBuffer
                                , ud_Address          := Address
                                , us_Length           := Size
                                );

    //no response
    if ( sd_retval <> 0 ) then
      LogError("@0286 (SafetyBaseFSoE::GetFSoEConnectionInfos) Config Read Error: Error reading routing info.");
      return;
    end_if;

    TempRoutingInfo := p_SDOResponseBuffer^.ud_Data$t_FSoERoutingInfoElement;

    // store the data in the connection info
    pActConnection^.SlaveAddress        := TempRoutingInfo.SlaveAddress;
    pActConnection^.MasterReadSize      := TempRoutingInfo.SafeOutputFrameSize;
    pActConnection^.MasterWriteSize     := TempRoutingInfo.SafeInputFrameSize;

    // the offset info depends on if we are master or slave
    if pActConnection^.Flags.IsMaster then
      pActConnection^.MasterReadOffset  := TempRoutingInfo.SafeOutputFrameOffset;
      pActConnection^.MasterWriteOffset := TempRoutingInfo.SafeInputFrameOffset;
    else
      pActConnection^.SlaveWriteOffset  := TempRoutingInfo.SafeOutputFrameOffset;
      pActConnection^.SlaveReadOffset   := TempRoutingInfo.SafeInputFrameOffset;
    end_if;

    pActConnection                  += sizeof(t_FSoEConnectionDetails);
    Address                         += Size;
  end_for;

//*****************************************************************************
//** CONNECTION INSTANCES                                                    **
//*****************************************************************************

  Address := SBF_SDO_ADDRESS_FSOE_CONN_INST;
  Size    := 4;

  //send request and receive data
  sd_retval := SDOReadCfgRequ ( p_SDORequestBuffer  := p_SDORequestBuffer
                              , p_SDOResponseBuffer := p_SDOResponseBuffer
                              , ud_Address          := Address
                              , us_Length           := Size
                              );

  //no response
  if ( sd_retval <> 0 ) then
    LogError("@0281 (SafetyBaseFSoE::GetFSoEConnectionInfos) Config Read Error: Error reading number of connections.");
    return;
  end_if;

  // check if it's the same number
  if ConnectionInfos.ConnectionNo <> p_SDOResponseBuffer^.ud_Data then
    LogError("@0287 (SafetyBaseFSoE::GetFSoEConnectionInfos) Config Read Error: Number of connections does not match (case 2).");
    return;
  end_if;

  Address += Size;

  pActConnection := ConnectionInfos.pFirstConnection;

  // get connection states
  for i := 0 to ConnectionInfos.ConnectionNo-1 do
    // get routing instance info of connections

    Size := 4;

    //send request and receive data
    sd_retval := SDOReadCfgRequ ( p_SDORequestBuffer  := p_SDORequestBuffer
                                , p_SDOResponseBuffer := p_SDOResponseBuffer
                                , ud_Address          := Address
                                , us_Length           := Size
                                );

    //no response
    if ( sd_retval <> 0 ) then
      LogError("@0288 (SafetyBaseFSoE::GetFSoEConnectionInfos) Config Read Error: Error reading size of routing instance info.");
      return;
    end_if;

    // calculate address of next connection (to check it later)
    NextAddress := Address + p_SDOResponseBuffer^.ud_Data;

    // get the flags
    Address   += Size;
    Size      := 4;

    //send request and receive data
    sd_retval := SDOReadCfgRequ ( p_SDORequestBuffer  := p_SDORequestBuffer
                                , p_SDOResponseBuffer := p_SDOResponseBuffer
                                , ud_Address          := Address
                                , us_Length           := Size
                                );

    //no response
    if ( sd_retval <> 0 ) then
      LogError("@0289 (SafetyBaseFSoE::GetFSoEConnectionInfos) Config Read Error: Error reading flags of routing instance info.");
      return;
    end_if;

    if ((p_SDOResponseBuffer^.ud_Data AND 1) <> 0) <> pActConnection^.Flags.IsMaster then
      LogError("@028A (SafetyBaseFSoE::GetFSoEConnectionInfos) Config Read Error: Master settings mismatch.");
      return;
    end_if;

    //! Flags
    //  Actually, type is 4 bytes in size but for compatibility reasons it is still used as 1 byte. As a result, bits 9-32 are currently not used.
    //  Bit1: 1, wenn FSoE-Master, 0=FSoE-Slave
    //  Bit2: 1, wenn die Slave-Adresse über den HW-Pfad ermittelt wird
    //  Bit3: 1, wenn CRC von der FW ermittelt werden muss
    //  Bit4: 1, wenn Interface und Slave
    //  Bit5: 1, wenn Multichannel verwendet werden, aber ein Multichannel ist nicht vorhanden und der Eingang auf 1 gesetzt wird.
    //  Bit6: 1, wenn der Adressvergabeservice verwendet werden soll
    //  Bit7: 1, wenn der Master beim Slave die Connection ID anfordert
    //  Bit8: 1, wenn es sich um ein HGW handelt
    //  Bit9: 1, wenn Assign Slave On Demand
    //  Bits 10-32: reserviert, sind auf 0 gesetzt und werden nicht ausgewertet

    //check size of FSoEFlags type --> possible are 1 or 4 byte
    pActConnection^.Flags := p_SDOResponseBuffer^.ud_Data$t_FSoEFlags;

    if (pActConnection^.Flags AND SM_FLAGS_FLEXCON_MASK) = SM_FLAGS_FLEXCON_NODE then
#ifdef SAFETY_DEBUG_LOGGING_ACTIVATED
      LogError(e_msg:="SafetyBaseFSoE: Found FSOE Connection of FlexConNode");
#endif
      sFlexCon.FoundNodeInConfig := TRUE;
    elsif (pActConnection^.Flags AND SM_FLAGS_FLEXCON_MASK) = SM_FLAGS_FLEXCON_HOST then
#ifdef SAFETY_DEBUG_LOGGING_ACTIVATED
      LogError(e_msg:="SafetyBaseFSoE: Found FSOE Connection of FlexConHost");
#endif
      sFlexCon.FoundHostInConfig := TRUE;
    end_if;

    // get the net size of the safe output data (only the bits for the I/Os without crc and stuff)
    Address   += Size;
    Size      := 2;

    //send request and receive data
    sd_retval := SDOReadCfgRequ ( p_SDORequestBuffer  := p_SDORequestBuffer
                                , p_SDOResponseBuffer := p_SDOResponseBuffer
                                , ud_Address          := Address
                                , us_Length           := Size
                                );

    //no response
    if ( sd_retval <> 0 ) then
      LogError("@028B (SafetyBaseFSoE::GetFSoEConnectionInfos) Config Read Error: Error reading safe output net size of routing instance info.");
      return;
    end_if;

    // we don't need the net size yet

    // get the net size of the safe input data (only the bits for the I/Os without crc and stuff)
    Address   += Size;
    Size      := 2;

    //send request and receive data
    sd_retval := SDOReadCfgRequ ( p_SDORequestBuffer  := p_SDORequestBuffer
                                , p_SDOResponseBuffer := p_SDOResponseBuffer
                                , ud_Address          := Address
                                , us_Length           := Size
                                );

    //no response
    if ( sd_retval <> 0 ) then
      LogError("@028C (SafetyBaseFSoE::GetFSoEConnectionInfos) Config Read Error: Error reading safe input net size of routing instance info.");
      return;
    end_if;

    // we don't need the net size yet

    // get the slave address
    Address   += Size;
    Size      := 2;

    //send request and receive data
    sd_retval := SDOReadCfgRequ ( p_SDORequestBuffer  := p_SDORequestBuffer
                                , p_SDOResponseBuffer := p_SDOResponseBuffer
                                , ud_Address          := Address
                                , us_Length           := Size
                                );

    //no response
    if ( sd_retval <> 0 ) then
      LogError("@028D (SafetyBaseFSoE::GetFSoEConnectionInfos) Config Read Error: Error reading slave address of routing instance info.");
      return;
    end_if;

    // the following settings are only available in the master
    if pActConnection^.Flags.IsMaster then

      // get the connection ID
      Address   += Size;
      Size      := 2;

      //send request and receive data
      sd_retval := SDOReadCfgRequ ( p_SDORequestBuffer  := p_SDORequestBuffer
                                  , p_SDOResponseBuffer := p_SDOResponseBuffer
                                  , ud_Address          := Address
                                  , us_Length           := Size
                                  );

      //no response
      if ( sd_retval <> 0 ) then
        LogError("@028E (SafetyBaseFSoE::GetFSoEConnectionInfos) Config Read Error: Error reading the connection ID of routing instance info.");
        return;
      end_if;

      pActConnection^.ConnectionID := p_SDOResponseBuffer^.ud_Data$UINT;

      // get transmission time
      Address   += Size;
      Size      := 2;

      //send request and receive data
      sd_retval := SDOReadCfgRequ ( p_SDORequestBuffer  := p_SDORequestBuffer
                                  , p_SDOResponseBuffer := p_SDOResponseBuffer
                                  , ud_Address          := Address
                                  , us_Length           := Size
                                  );

      //no response
      if ( sd_retval <> 0 ) then
        LogError("@028F (SafetyBaseFSoE::GetFSoEConnectionInfos) Config Read Error: Error reading the transmission time of routing instance info.");
        return;
      end_if;

      pActConnection^.TransmissionTime_ms := p_SDOResponseBuffer^.ud_Data$UINT;

      // get length of communication parameters (must be 2)
      Address   += Size;
      Size      := 2;

      //send request and receive data
      sd_retval := SDOReadCfgRequ ( p_SDORequestBuffer  := p_SDORequestBuffer
                                  , p_SDOResponseBuffer := p_SDOResponseBuffer
                                  , ud_Address          := Address
                                  , us_Length           := Size
                                  );

      //no response
      if ( sd_retval <> 0 ) then
        LogError("@0290 (SafetyBaseFSoE::GetFSoEConnectionInfos) Config Read Error: Error reading the length of the communication parameters of routing instance info.");
        return;
      end_if;

      if p_SDOResponseBuffer^.ud_Data$UINT <> 2 then
        LogError("@0291 (SafetyBaseFSoE::GetFSoEConnectionInfos) Config Read Error: Length of communication parameters is wrong.");
        return;
      end_if;

      // skip FSoE watchdog time in ms
      Address   += Size;
      Size      := 2;

      // get size of application parameters
      Address   += Size;
      Size      := 2;

      //send request and receive data
      sd_retval := SDOReadCfgRequ ( p_SDORequestBuffer  := p_SDORequestBuffer
                                  , p_SDOResponseBuffer := p_SDOResponseBuffer
                                  , ud_Address          := Address
                                  , us_Length           := Size
                                  );

      //no response
      if ( sd_retval <> 0 ) then
        LogError("@0292 (SafetyBaseFSoE::GetFSoEConnectionInfos) Config Read Error: Error reading the length of the application parameters of routing instance info.");
        return;
      end_if;

      // skip length
      Address   += Size;

      // skip application parameters
      Size      := p_SDOResponseBuffer^.ud_Data$USINT;
      Address   += Size;

      // get to a 4 byte aligned address
      if (Address MOD 4) then
        Address := Address + (4 - (Address MOD 4)); //increase memory, up to a value, which could be divided by 4
      end_if;

      // get size of hw path
      Size      := 4;

      //send request and receive data
      sd_retval := SDOReadCfgRequ ( p_SDORequestBuffer  := p_SDORequestBuffer
                                  , p_SDOResponseBuffer := p_SDOResponseBuffer
                                  , ud_Address          := Address
                                  , us_Length           := Size
                                  );

      //no response
      if ( sd_retval <> 0 ) then
        LogError("@0293 (SafetyBaseFSoE::GetFSoEConnectionInfos) Config Read Error: Error reading the hardware path length of routing instance info.");
        return;
      end_if;

      // get the hardware path
      Address   += Size;
      Size      := p_SDOResponseBuffer^.ud_Data$USINT;

      if Size = 0 then
        LogError("@0294 (SafetyBaseFSoE::GetFSoEConnectionInfos) Config Read Error: Hardware path length is zero.");
        return;
      end_if;

      //send request and receive data
      sd_retval := SDOReadCfgRequ ( p_SDORequestBuffer  := p_SDORequestBuffer
                                  , p_SDOResponseBuffer := p_SDOResponseBuffer
                                  , ud_Address          := Address
                                  , us_Length           := Size
                                  );

      //no response
      if ( sd_retval <> 0 ) then
        LogError("@0295 (SafetyBaseFSoE::GetFSoEConnectionInfos) Config Read Error: Error reading the hardware path of routing instance info.");
        return;
      end_if;

      // save hardware path into structure
      pActConnection^.SlavePathLen      := Size;
      pActConnection^.pSlavePath$pVoid  := ToStdLib.Malloc(size:=Size);

      if pActConnection^.pSlavePath = NIL then
        LogError("@0296 (SafetyBaseFSoE::GetFSoEConnectionInfos) Failed to allocate memory for the slave hardware path at the routing instance info.");
        return;
      end_if;

      _memcpy(ptr1:=pActConnection^.pSlavePath, ptr2:=#p_SDOResponseBuffer^.ud_Data, cntr:=pActConnection^.SlavePathLen);

      Address         += Size;

      // get to a 4 byte aligned address
      if (Address MOD 4) then
        Address := Address + (4 - (Address MOD 4)); //increase memory, up to a value, which could be divided by 4
      end_if;

      // get size of compressed hw path
      Size      := 4;

      //send request and receive data
      sd_retval := SDOReadCfgRequ ( p_SDORequestBuffer  := p_SDORequestBuffer
                                  , p_SDOResponseBuffer := p_SDOResponseBuffer
                                  , ud_Address          := Address
                                  , us_Length           := Size
                                  );

      //no response
      if ( sd_retval <> 0 ) then
        LogError("@0297 (SafetyBaseFSoE::GetFSoEConnectionInfos) Config Read Error: Error reading the compressed hardware path length of routing instance info.");
        return;
      end_if;

      // get the hardware path
      Address   += Size;
      Size      := p_SDOResponseBuffer^.ud_Data$USINT;

      //send request and receive data
      sd_retval := SDOReadCfgRequ ( p_SDORequestBuffer  := p_SDORequestBuffer
                                  , p_SDOResponseBuffer := p_SDOResponseBuffer
                                  , ud_Address          := Address
                                  , us_Length           := Size
                                  );

      //no response
      if ( sd_retval <> 0 ) then
        LogError("@0298 (SafetyBaseFSoE::GetFSoEConnectionInfos) Config Read Error: Error reading the compressed hardware path of routing instance info.");
        return;
      end_if;

      // save compressed hardware path into structure
      pActConnection^.SlavePathCompLen      := Size;
      pActConnection^.pSlavePathComp$pVoid  := ToStdLib.Malloc(size:=Size);

      if pActConnection^.pSlavePathComp = NIL then
        LogError("@0299 (SafetyBaseFSoE::GetFSoEConnectionInfos) Failed to allocate memory for the compressed slave hardware path at the routing instance info.");
        return;
      end_if;

      _memcpy(ptr1:=pActConnection^.pSlavePathComp, ptr2:=#p_SDOResponseBuffer^.ud_Data, cntr:=pActConnection^.SlavePathCompLen);

      if  (pActConnection^.pSlavePathComp^ = 6) &
          ((pActConnection^.pSlavePathComp + 5)^$HDINT AND 16#00FFFFFF) = 0 then

        // special IP: (0.0.0.x)
        // if custom ip is detected change pathcomp type from 6 (IP) to 3 (Interface)
        pActConnection^.pSlavePathComp^ :=3;
      end_if;

      //Get slot ID and communication ID from HGW
      if pActConnection^.Flags.IsHGW then

        //Get machinenumber of FUB
        sd_retval := SDOReadCfgRequ ( p_SDORequestBuffer  := p_SDORequestBuffer
                                    , p_SDOResponseBuffer := p_SDOResponseBuffer
                                    , ud_Address          := SBF_SDO_ADDRESS_HGW_FUB_BASE_ADDRESS + SBF_SDO_ADDRESS_HGW_OFFSET_MACHINENUMBER
                                    , us_Length           := 4
                                    , b_UseCache          := FALSE
                                    );

        //no response
        if ( sd_retval <> 0 ) then
          LogError("@03DA (SafetyBaseFSoE::GetFSoEConnectionInfos) Config Read Error: Error reading the machinenumber of routing instance info.");
          return;
        end_if;

        sHGW.udMachineNrb := p_SDOResponseBuffer^.ud_Data$UDINT;

        // get the Slot ID
        Address   += Size;
        Size      := 2;

        //send request and receive data
        sd_retval := SDOReadCfgRequ ( p_SDORequestBuffer  := p_SDORequestBuffer
                                    , p_SDOResponseBuffer := p_SDOResponseBuffer
                                    , ud_Address          := Address
                                    , us_Length           := Size
                                    );

        //no response
        if ( sd_retval <> 0 ) then
          LogError("@03DB (SafetyBaseFSoE::GetFSoEConnectionInfos) Config Read Error: Error reading the communication ID of routing instance info.");
          return;
        end_if;

        sHGW.uiCommunicationID := p_SDOResponseBuffer^.ud_Data$UINT;

        // get the communication ID
        Address   += Size;
        Size      := 2;

        //send request and receive data
        sd_retval := SDOReadCfgRequ ( p_SDORequestBuffer  := p_SDORequestBuffer
                                    , p_SDOResponseBuffer := p_SDOResponseBuffer
                                    , ud_Address          := Address
                                    , us_Length           := Size
                                    );

        //no response
        if ( sd_retval <> 0 ) then
          LogError("@03DC (SafetyBaseFSoE::GetFSoEConnectionInfos) Config Read Error: Error reading the slot ID of routing instance info.");
          return;
        end_if;

        sHGW.uiSlotID := p_SDOResponseBuffer^.ud_Data$UINT;

        //save fsoe pdo offsets and length
        sHGW.InputPDOLength  := pActConnection^.MasterWriteSize;
        sHGW.OutputPDOLength := pActConnection^.MasterReadSize;
        if pActConnection^.Flags.IsMaster then
          sHGW.InputPDOOffset  := pActConnection^.MasterWriteOffset;
          sHGW.OutputPDOOffset := pActConnection^.MasterReadOffset;
        else
          sHGW.InputPDOOffset  := pActConnection^.SlaveWriteOffset;
          sHGW.OutputPDOOffset := pActConnection^.SlaveReadOffset;
        end_if;
        sHGW.uiTransmissionTime_ms := pActConnection^.TransmissionTime_ms;
      end_if;

      Address         += Size;

      // get to a 4 byte aligned address
      if (Address MOD 4) then
        Address := Address + (4 - (Address MOD 4)); //increase memory, up to a value, which could be divided by 4
      end_if;

      if Address > NextAddress then
        LogError("@029A (SafetyBaseFSoE::GetFSoEConnectionInfos) Config Read Error: Structure size mismatch.");
        return;
      end_if;
    end_if;

    Address         := NextAddress;
    pActConnection  += sizeof(t_FSoEConnectionDetails);
  end_for;

END_FUNCTION

FUNCTION SafetyBaseFSoE::FreeFSoEConnectionInfos
  VAR
    i               : UDINT;
    pActConnection  : ^t_FSoEConnectionDetails;
  END_VAR

  if (ConnectionInfos.ConnectionNo = 0) | (ConnectionInfos.pFirstConnection = NIL) then
    // nothing to free
    return;
  end_if;

  // check if all connections have been initialized
  pActConnection := ConnectionInfos.pFirstConnection;
  for i := 0 to ConnectionInfos.ConnectionNo-1 do
    if pActConnection^.ConnectionState = FCS_NOT_INITIALIZED then
      // not yet time to free them
      return;
    end_if;

    pActConnection += sizeof(t_FSoEConnectionDetails);
  end_for;

  pActConnection := ConnectionInfos.pFirstConnection;
  for i := 0 to ConnectionInfos.ConnectionNo-1 do
    // free hardware path memory

    if pActConnection^.pSlavePath then
      ToStdLib.Free(mptr:=pActConnection^.pSlavePath);
    end_if;

    if pActConnection^.pSlavePathComp then
      ToStdLib.Free(mptr:=pActConnection^.pSlavePathComp);
    end_if;

    pActConnection += sizeof(t_FSoEConnectionDetails);
  end_for;

  // free the connectionlist
  ToStdLib.Free(mptr:=ConnectionInfos.pFirstConnection);
  ConnectionInfos.pFirstConnection := NIL;
  ConnectionInfos.ConnectionNo := 0;

END_FUNCTION

FUNCTION SafetyBaseFSoE::CheckFSoEConnections
  VAR
    MyPara 	            : CmdStruct;
    MyResult	          : results;
    i                   : UDINT;
    pActConnection      : ^t_FSoEConnectionDetails;
    SDORequestBuffer    : SDORequReadConfig;
    SDOResponseBuffer   : ARRAY [0..SBF_SDO_MAX_LENGTH-1] OF USINT;
    p_SDORequestBuffer 	: ^SDORequReadConfig;
    p_SDOResponseBuffer : ^SDORespReadConfig;
    UnInifializedNo     : UDINT;
    sd_retval           : DINT;
  END_VAR

  // there were some of the FSoE connections not initialized when fetching the configuration data => update them

  UnInifializedNo := 0;

  //SDO request for this command has 5 bytes additional to the header
  p_SDORequestBuffer := #SDORequestBuffer;

  //SDO response for this command can have maximum additional data
  p_SDOResponseBuffer := (#SDOResponseBuffer)$^SDORespReadConfig;

  //calculate length without crc
  p_SDORequestBuffer^.StdHeader.Len := sizeof(SDORequReadConfig) - sizeof(SDOHeader.StdHeader.CRC);

  //type
  p_SDORequestBuffer^.StdHeader.Typ := SDO_STD;

  //command for reading config data
  p_SDORequestBuffer^.StdHeader.Cmd := SBF_SDO_COMMAND_READ;

  // reset cache, because it may contain an old access on the same address => we want fresh data
  CachedSize := 0;

  pActConnection := ConnectionInfos.pFirstConnection;

  for i := 0 to ConnectionInfos.ConnectionNo-1 do
    if pActConnection^.ConnectionState = FCS_NOT_INITIALIZED then
      UnInifializedNo += 1;

      //send request and receive data
      sd_retval := SDOReadCfgRequ ( p_SDORequestBuffer  := p_SDORequestBuffer
                                  , p_SDOResponseBuffer := p_SDOResponseBuffer
                                  , ud_Address          := SBF_SDO_ADDRESS_FSOE_CONN_STATE + 2 + i
                                  , us_Length           := 1
                                  );

      //no response
      if ( sd_retval <> 0 ) then
        LogError("@0283 (SafetyBaseFSoE::CheckFSoEConnections) Config Read Error: Error reading connection state.");
        return;
      end_if;

      // get connection state
      pActConnection^.ConnectionState := (p_SDOResponseBuffer^.ud_Data$USINT AND 2#0111)$t_FSoEConnectionState;

      if pActConnection^.ConnectionState <> FCS_NOT_INITIALIZED then
        UnInifializedNo -= 1;

        // get the corresponding slave address number

        //send request and receive data
        sd_retval := SDOReadCfgRequ ( p_SDORequestBuffer  := p_SDORequestBuffer
                                    , p_SDOResponseBuffer := p_SDOResponseBuffer
                                    , ud_Address          := SBF_SDO_ADDRESS_FSOE_ROUTING_INFO + 2 + i * sizeof(t_FSoERoutingInfoElement)
                                    , us_Length           := sizeof(t_FSoERoutingInfoElement)
                                    );

        //no response
        if ( sd_retval <> 0 ) then
          LogError("@0286 (SafetyBaseFSoE::CheckFSoEConnections) Config Read Error: Error reading routing info.");
          return;
        end_if;

        pActConnection^.SlaveAddress := p_SDOResponseBuffer^.ud_Data$t_FSoERoutingInfoElement.SlaveAddress;

        if pActConnection^.SlaveAddress = 0 then
          LogError("@029B (SafetyBaseFSoE::CheckFSoEConnections) Connection initialized but slave address is still zero!");
        end_if;
      end_if;
    end_if;

    pActConnection                  += sizeof(t_FSoEConnectionDetails);
  end_for;

  // if all connections are initialized => tell the safety manager
  if (UnInifializedNo = 0) & pSafetyManagerThis then
    MyPara.uiCmd    := CMD_SM_FSOE_CON_INITIALIZED;
    MyPara.aPara[0] := SafetyNumber$DINT;
    MyPara.aPara[1] := ConnectionInfos.ConnectionNo$DINT;
    MyPara.aPara[2] := ConnectionInfos.pFirstConnection$DINT;

    if pSafetyManagerThis^.NewInst(#MyPara, #MyResult) = READY then
      // we don't need this memory anymore
      FreeFSoEConnectionInfos();
    end_if;
  end_if;

END_FUNCTION

FUNCTION VIRTUAL GLOBAL SafetyBaseFSoE::GetDiagConnect::NewInst
  VAR_INPUT
    pPara 	: ^CmdStruct;
    pResult 	: ^Results;
  END_VAR
  VAR_OUTPUT
    ret_code 	: IprStates;
  END_VAR

  ret_code := READY;

  CASE pPara^.uiCmd OF

    CMD_SM_DIAG_GET_INFO:

      //Subcommand
      case pPara^.aPara[0] of
//*****************************************************************************
        SBCMD_SM_DIAG_GET_INFO:
          pResult^.aData[0] :=  GetDiagInfo(pDiagInfo:=(pPara^.aPara[1])$^SafetyDiagInfo);

//*****************************************************************************
        SBCMD_SM_DIAG_GET_STATE:
          pResult^.aData[0] :=  GetDiagState(pDiagState:=(pPara^.aPara[1])$^SafetyDiagState);

//*****************************************************************************
        SBCMD_SM_DIAG_FETCH_INFO:
      //Fetch Diag Info for uCx
          FetchDiagInfo(ucChoice:=pPara^.aPara[1]$USINT);

//*****************************************************************************
        SBCMD_SM_DIAG_FETCH_STATE:
          FetchDiagState();

//*****************************************************************************
        SBCMD_SM_DIAG_IS_SAVE_LOG_ACTIVE:
          pResult^.aData[0] := SaveLogActive();

//*****************************************************************************
        SBCMD_SM_DIAG_SAVE_LOGFILE:
          pResult^.aData[0] := (SaveLog(ucChoice:=(pPara^.aPara[1])$USINT, pDPNE:=(pPara^.aPara[2])$^CHAR))$USINT;

//*****************************************************************************
        SBCMD_SM_DIAG_GET_SAVE_LOGFILE_STATE:
          pResult^.aData[0] := DiagVars.SavingLogSuccessful$USINT;

//*****************************************************************************
        SBCMD_SM_DIAG_GET_SAFETY_NUMBER:
          pResult^.aData[0]$UDINT := SafetyNumber;

//*****************************************************************************
        SBCMD_SM_DIAG_GET_SAFETY_STATE:
          pResult^.aData[0] := SafetyState$USINT;

//*****************************************************************************
        SBCMD_SM_DIAG_IS_DIAGNOSE_AVAILABLE:
          pResult^.aData[0] := TRUE;

//*****************************************************************************
        SBCMD_SM_DIAG_GET_CHANNEL_INFO:
          pResult^.aData[0] := GetChannelInfo(pErrorMemUser:=(pPara^.aPara[1])$^UINT, pErrorMem:=#aErrorMem[1], ErrorDataLength:=aErrorMem[0] - 1);
          pResult^.aData[1] := aErrorMem[0] - 1;

//*****************************************************************************
        SBCMD_SM_DIAG_FETCH_CHANNEL_INFO:
          FetchChannelInfo();

      END_CASE;
    else
      TRACE("(SafetyBaseFSoE::GetDiagConnect::NewInst) Unknown command!");
      ret_code := ERROR;
  END_CASE;

END_FUNCTION

FUNCTION SafetyBaseFSoE::GetNewMemSize
  VAR_INPUT
    Required 	: UDINT;
  END_VAR
  VAR_OUTPUT
    NextBiggerBlockSize 	: UDINT;
  END_VAR

  // how many complete blocks are necessary
  NextBiggerBlockSize := Required / SBF_CONFIG_MEMORY_BLOCK_SIZE;

  // is there also an incomplete block?
  if Required MOD SBF_CONFIG_MEMORY_BLOCK_SIZE then
    NextBiggerBlockSize += 1;
  end_if;

  // now that we have the number of blocks necessary => get number of bytes
  NextBiggerBlockSize *= SBF_CONFIG_MEMORY_BLOCK_SIZE;

END_FUNCTION

FUNCTION SafetyBaseFSoE::CheckAddDynSlaveResponse
  VAR_INPUT
    pAddDynSlaveRsp 	: ^t_AddDynSlaveResponse;
  END_VAR
  VAR_OUTPUT
    ResponseOk 	: BOOL;
  END_VAR

  // check if any of the offset/length combination exceeds our access to the module
  if ((pAddDynSlaveRsp^.OffsetSafeInData  + pAddDynSlaveRsp^.LenSafeInData ) > MyPDOWriteSize) |
     ((pAddDynSlaveRsp^.OffsetSafeOutData + pAddDynSlaveRsp^.LenSafeOutData) > MyPDOReadSize ) then
    ResponseOk := FALSE;

    LogError("@029C (SafetyBaseFSoE::CheckAddDynSlaveResponse) Invalid offset/length combination of read or write data in AddDynSlave response.");
  else
    ResponseOk := TRUE;
  end_if;

END_FUNCTION

FUNCTION SafetyBaseFSoE::GetChannelInfo
  VAR_INPUT
    pErrorMemUser 	: ^UINT;
    pErrorMem 	: ^USINT;
    ErrorDataLength 	: INT;
  END_VAR
  VAR_OUTPUT
    StateReady 	: BOOL;
  END_VAR
  VAR
    i   : INT;
  END_VAR

  StateReady := DiagVars.UserErrorInfoReady;

  if StateReady then
    //copy error values in UserArray
    for i := 0 to ErrorDataLength-1 do

      pErrorMemUser^ := pErrorMem^;

      //Add 1000 to each errorvalue so that it matches the value in SafetyDesigner.
      if (pErrorMemUser^ <> 0) then
        pErrorMemUser^ += 1000;
      end_if;

      //set pointer to next entry
      pErrorMemUser += sizeof(UINT);
      pErrorMem += sizeof(USINT);
    end_for;
  end_if;

END_FUNCTION

FUNCTION VIRTUAL GLOBAL SafetyBaseFSoE::FetchChannelInfo

  DiagVars.UserErrorInfoReady := FALSE;
  DiagVars.UserWantsErrorInfo := TRUE;

END_FUNCTION

#pragma warning(disable:73);
FUNCTION VIRTUAL SafetyBaseFSoE::SafeActModuleConfig
  VAR_INPUT
    sActModuleConfig 	: t_ModuleCfg;
  END_VAR
  //overwrite this function at derived class to safe module config
END_FUNCTION
#pragma warning(default:73);
